// TIA Portal V21 export
// export: Created 2026-11-22T02:34:16.8188654Z, ExportSetting WithDefaults, DisplayName Totally Integrated Automation Portal, DisplayVersion V21 Update 3, DisplayName STEP 7 Professional, DisplayVersion V21 Update 3, DisplayName STEP 7 Safety, DisplayVersion V21, DisplayName Tech WebApplication, DisplayVersion V21, DisplayName WinCC Basic/Comfort/Advanced, DisplayVersion V21 Update 3, DisplayName WinCC Unified, DisplayVersion V21 Update 3
Screen "D_Bar_2"  800x480, Number=466
  ScreenLayer "Layer_0"
    Bar "PV_Pct_0_100" at 6,4 size 40x120  CountSubDivisions=5, IntegerDigits=3, LargeTickLabelingStep=1, MaximumValue=100, Precision=2, StyleItem=Bar
      ProcessValue := D_Pct
    TextField "Label_PV_Pct_0_100" at 6,156 size 88x16  StyleItem=Text field, Text="PV_Pct_0_100"
    Bar "PV_Pct_MaxMin" at 98,4 size 40x120  CountSubDivisions=5, IntegerDigits=3, LargeTickLabelingStep=1, MaximumValue=5, MinimumValue=-5, Precision=2, StyleItem=Bar
      ProcessValue := D_Pct
      MaximumValue := D_Max
      MinimumValue := D_Min
    TextField "Label_PV_Pct_MaxMin" at 98,156 size 88x16  StyleItem=Text field, Text="PV_Pct_MaxMin"
    IOField "State" at 4,454 size 60x22  DataFormat=Decimal, FormatPattern=9, Mode=Output, StyleItem=I/O field
      ProcessValue := D_State
    Button "S1" at 70,454 size 40x22  Mode=Text, StyleItem=Button, TextOff="S1", TextOn="S1"
      on Click: SetS1()
    Button "S2" at 114,454 size 40x22  Mode=Text, StyleItem=Button, TextOff="S2", TextOn="S2"
      on Click: SetS2()
    Button "S3" at 158,454 size 40x22  Mode=Text, StyleItem=Button, TextOff="S3", TextOn="S3"
      on Click: SetS3()
    Button "S4" at 202,454 size 40x22  Mode=Text, StyleItem=Button, TextOff="S4", TextOn="S4"
      on Click: SetS4()
    Button "Next" at 756,454 size 40x22  Mode=Text, StyleItem=Button, TextOff="Next", TextOn="Next"
      on Click: ActivateScreen(Screen name := D_Switch_1, Object number := 0)
